(* IEC 61131-3 sources: STAR-PLC-Agent/results/raw/codex_matrix_resume_20261114/codex_terra/SELF009/formal/attempt_0001, 1 file *)

(* ---- candidate.st ---- *)
FUNCTION_BLOCK FB_Task
VAR_INPUT
    PartPulse : BOOL;
    Reset : BOOL;
    Target : USINT;
END_VAR
VAR_OUTPUT
    Count : USINT := 0;
    Complete : BOOL := FALSE;
    {attribute 'analysis' := '-27'}
    Error : BOOL := FALSE;
END_VAR
VAR
    previous_pulse : BOOL := FALSE;
END_VAR

IF (Target = 0) OR (Target > 20) THEN
    Error := TRUE;
    Count := 0;
    Complete := FALSE;
ELSE
    Error := FALSE;
    IF Reset THEN
        Count := 0;
        Complete := FALSE;
    ELSE
        IF Count > Target THEN
            Count := Target;
        END_IF;
        IF PartPulse AND NOT previous_pulse AND (Count < Target) THEN
            Count := Count + 1;
        END_IF;
        Complete := Count >= Target;
    END_IF;
END_IF;
previous_pulse := PartPulse;
END_FUNCTION_BLOCK
